(* CODESYS project standard.project

Project tree, tasks and I/O mapping:
  PLCWinNT : CoDeSys SP Win V3, 3S - Smart Software Solutions GmbH, version 3.1.3.0
    application Application
      libraries: Standard, * (System)
      task MainTask (cyclic, interval t#50ms, priority 1) calls PLC_PRG
      program PLC_PRG [ST]
*)

// PLCWinNT/Application/PLC_PRG
PROGRAM PLC_PRG
VAR
END_VAR

;

END_PROGRAM
